Fanuc KAREL source: kt00445.KL

-- PROVISIONAL review KL for V1013-1; original PC SHA256 424463f83a9380557e6aa7d8cf840462eea0def1b2250981698f72cf1dbf0f75
-- Incomplete behavior may be omitted. Consult companion uncertainty JSON. Do not deploy.
PROGRAM KT00445
%NOLOCKGROUP
VAR
  B1 : BOOLEAN
  B2 : BOOLEAN
  OUT : BOOLEAN
BEGIN
  -- UNRESOLVED_PC offsets 5-12; opcodes 9D,23
  -- UNRESOLVED_PC offsets 17-24; opcodes 9C,23
  -- UNRESOLVED_PC offsets 29-36; opcodes 9D,23
  -- UNRESOLVED_PC offsets 41-48; opcodes 9C,23
  -- UNRESOLVED_PC offsets 53-72; opcodes 21,21,5C,23
  -- UNRESOLVED_PC offsets 77-81; opcodes 7F
END KT00445
